// Simulation program for the Valve Characterization sample.
// Models a non-linear hydraulic valve: integrates the (non-linear) spool velocity to an actual
// position and feeds simulated I/O, so the sample runs without real hardware.
PROGRAM Simu
VAR
	ActPos AT%Q*:	DINT;
	SetVelo AT%I*:	INT;
	PressureA AT%Q*:	INT;
 
 	fSetVelo:	LREAL;
 	fActPos:	LREAL;

	fSetVeloNonLinear: LREAL;
END_VAR


fSetVelo:=INT_TO_LREAL(SetVelo)/32767*500.0;

IF fSetVelo > 0.0 THEN
	fSetVeloNonLinear := (1-COS(fSetVelo/500.0*3.14))/2.0*500.0;
ELSE
	fSetVeloNonLinear := -(1-COS(fSetVelo/500.0*3.14))/2.0*500.0;
END_IF
//fSetVeloNonLinear:=fSetVelo;
fActPos:=fActPos+fSetVeloNonLinear*0.002;

fActPos:=MIN(MAX(fActPos,0.0),500.0);
ActPos:=LREAL_TO_DINT(fActPos * 1000.0);

END_PROGRAM

(* stored: Version 1.1.0.1, ProductVersion 3.1.4026.4
   POU Simu: Id {bc1941f6-7ebc-436a-b9d8-839f2afffadf}, SpecialFunc None *)
